// TIA Portal V18 export
TYPE "Udt_Data_AGVToScala"
   STRUCT
      POPID : String[10];   // POPID
      CU : String[10];   // CU
      AGVNumber : Int;   // Número AGV
      ProductOK : Bool;   // Produto recebido OK
      ProductNOK : Bool;   // Falha produto recebido Scala
      AGVRedCard : Bool;   // AGV com trabalho
      Spare4 : Bool;   // Reserva
      Spare5 : Bool;   // Reserva
      Spare6 : Bool;   // Reserva
      Spare7 : Bool;   // Reserva
      Spare8 : Bool;   // Reserva
      Spare9 : Bool;   // Reserva
      Spare10 : Bool;   // Reserva
      Spare11 : Bool;   // Reserva
      Spare12 : Bool;   // Reserva
      Spare13 : Bool;   // Reserva
      Spare14 : Bool;   // Reserva
      Spare15 : Bool;   // Reserva
      Spare16 : Bool;   // Reserva
   END_STRUCT;
END_TYPE
